// TIA Portal project "Texts" (V21)

(* hardware
DEVICE "PLC_Texts"  S7-1500 station
   slot 0: "Rail_0"  Rack  6ES7 590-1***0-0AA0
   slot 1: "PLC_Texts"  CPU 1516-3 PN/DP  6ES7 516-3AN02-0AB0  V2.9
      slot 3: "CPU display_1"  6ES7591-1BA00-0AA0
      slot 32768: "PROFINET interface_1"  X1
         slot 32769: "Port_1"  X1 P1
         slot 32770: "Port_2"  X1 P2
      slot 33024: "PROFINET interface_2"  X2
         slot 33025: "Port_1"  X2 P1
      slot 33280: "DP interface_1"  X3
      slot 34817: "Virtual CP interface port_1"  Virtual CP interface port  Virtual CP interface port
*)

// ===== PLC "PLC_Texts"  CPU 1516-3 PN/DP =====
// protected blocks, not shown: "Sealed"

VAR_GLOBAL   // PLC tag table "Signals"
   "levelSensor" AT %IW10 : Int;   // Füllstandsensor / Level sensor / Capteur de niveau
   "pumpOn" AT %Q4.0 : Bool;   // Pumpe ein / Pump on / Pompe en marche
   "spare" AT %Q4.1 : Bool;   // Spare output
END_VAR

DATA_BLOCK "TankA"   // DB1
{ S7_Optimized_Access := 'TRUE' }
VERSION : 0.1
// stored: InstanceOfName Tank
"Tank"
BEGIN
END_DATA_BLOCK

DATA_BLOCK "TankB"   // DB2
{ S7_Optimized_Access := 'TRUE' }
VERSION : 0.1
// stored: InstanceOfName Tank
"Tank"
BEGIN
END_DATA_BLOCK

DATA_BLOCK "Recipe"   // DB30
TITLE = Rezept / Recipe / Recette
{ S7_Optimized_Access := 'TRUE' }
// Werte des Rezepts / Values of the recipe / Valeurs de la recette
   VAR
      target : Int := 500;   // Sollfüllstand in mm / Target level in mm / Niveau de consigne en mm
      hysteresis : Int := 20;   // Hysteresis in mm
   END_VAR
BEGIN
END_DATA_BLOCK

// folder: Closed

DATA_BLOCK "SealedA"   // DB3
{ S7_Optimized_Access := 'TRUE' }
VERSION : 0.1
// stored: InstanceOfName Sealed
"Sealed"
BEGIN
END_DATA_BLOCK

// folder: (top level)

FUNCTION_BLOCK "Tank"   // FB1, SCL
TITLE = Behälter überwachen / Watch the tank / Surveiller le réservoir
{ S7_Optimized_Access := 'TRUE' }
VERSION : 0.1
// Meldet einen hohen und einen niedrigen Füllstand. / Reports a high and a low level. / Signale un niveau haut et un niveau bas.
   VAR_INPUT
      level : Int;   // Füllstand in mm
      high : Bool;   // Grenzwert oben erreicht
      low : Bool;
      state : Int;   // Zustand, Index in die Textliste States
   END_VAR
   VAR
      highAlarm : Program_Alarm;
      lowAlarm : Program_Alarm;
   END_VAR
BEGIN

    #highAlarm(SIG := #high, SD_1 := #level);
    #lowAlarm(SIG := #low, SD_1 := #level, SD_2 := #state);
END_FUNCTION_BLOCK

FUNCTION_BLOCK "Valve"   // FB20, LAD
TITLE = Ventil / Valve / Vanne
{ S7_Optimized_Access := 'TRUE' }
// Ein Ventil mit Rückmeldung. / A valve with feedback. / Une vanne avec retour d'information.
   VAR_INPUT
      open : Bool;   // Ventil öffnen / Open the valve / Ouvrir la vanne
      close : Bool;   // Close the valve
   END_VAR
   VAR_OUTPUT
      opened : Bool;   // Vanne ouverte
   END_VAR
   VAR
      moving : Bool;   // Ventil fährt / Valve is moving / La vanne se déplace
   END_VAR
BEGIN

REGION Network 1: Öffnen / Open / Ouvrir
   // Öffnen setzt das Fahren. / Opening starts the travel. / L'ouverture lance le déplacement.
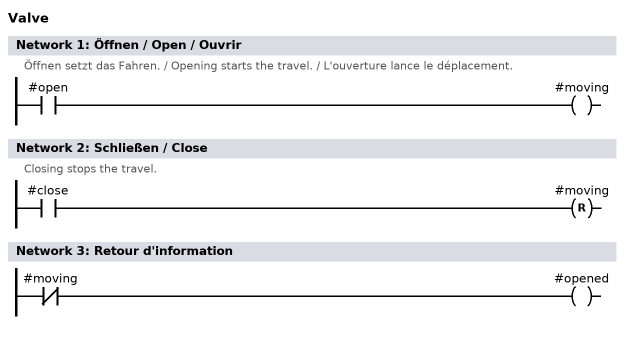
   RUNG wire#powerrail
      Contact( #open )
      Coil( #moving )
   END_RUNG
   // the same network as SCL:
   #moving := #open;
END_REGION

REGION Network 2: Schließen / Close
   // Closing stops the travel.
   RUNG wire#powerrail
      Contact( #close )
      R_Coil( #moving )
   END_RUNG
   // the same network as SCL:
   IF #close THEN #moving := FALSE; END_IF;
END_REGION

REGION Network 3: Retour d'information
   RUNG wire#powerrail
      I_Contact( #moving )
      Coil( #opened )
   END_RUNG
   // the same network as SCL:
   #opened := NOT #moving;
END_REGION
END_FUNCTION_BLOCK